// TIA Portal V20 export
FUNCTION_BLOCK "OM_PRM_Access"   // FB82, LAD
{ S7_Optimized_Access := 'TRUE' }
// stored: MemoryReserve 100, SetENOAutomatically false
   VAR_INPUT
      Inputdata_RW_Drv2PLC : "AZ_PrmRW_Drv2PLC";
      ReadParameterID : Word;
      WriteParameterID : Word;
      WriteData : DWord;
      "WR-REQ" : Bool;
   END_VAR
   VAR_OUTPUT
      Outputdata_RW_PLC2Drv : "AZ_PrmRW_PLC2Drv";
      ReadParameterID_R : Word;
      WriteParameterID_R : Word;
      ReadData : DWord;
      "WR-SET-ERR" : Bool;
      "WR-IF-ERR" : Bool;
      "WR-NV-ERR" : Bool;
      "WR-EXE-ERR" : Bool;
      "WR-ERR" : Bool;
      "RD-ERR" : Bool;
      "WR-END" : Bool;
      "SYS-BSY" : Bool;
   END_VAR
BEGIN

REGION Network 1
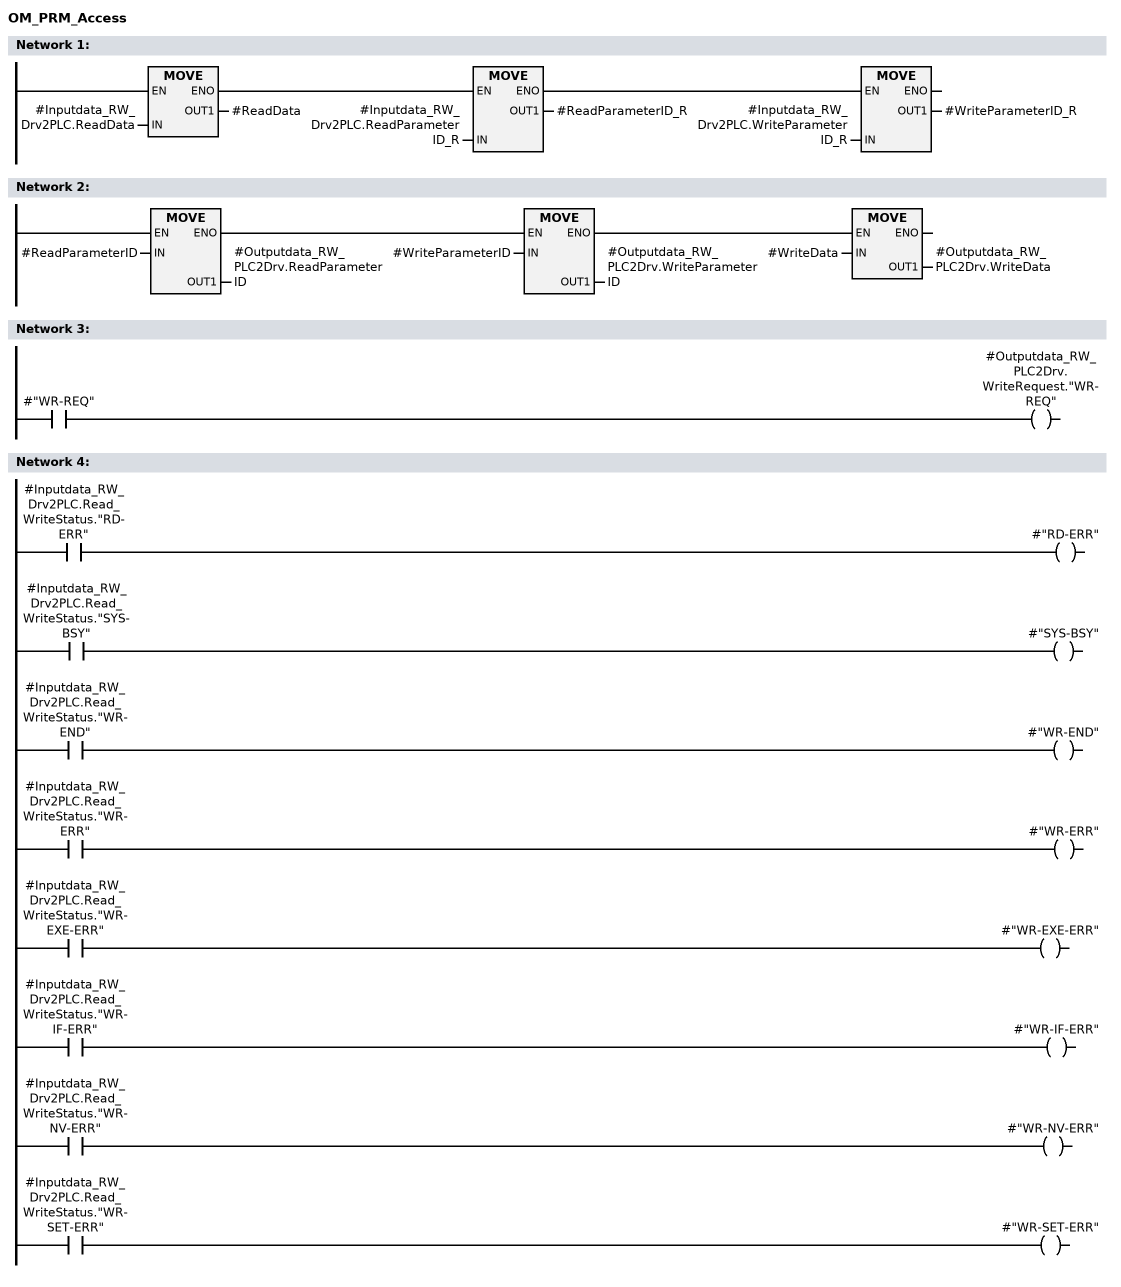
   RUNG wire#powerrail
      Move(in := #Inputdata_RW_Drv2PLC.ReadData, out1 => #ReadData)
      Move(in := #Inputdata_RW_Drv2PLC.ReadParameterID_R, out1 => #ReadParameterID_R)
      Move(in := #Inputdata_RW_Drv2PLC.WriteParameterID_R, out1 => #WriteParameterID_R)
   END_RUNG
   // the same network as SCL:
   #ReadData := #Inputdata_RW_Drv2PLC.ReadData;
   #ReadParameterID_R := #Inputdata_RW_Drv2PLC.ReadParameterID_R;
   #WriteParameterID_R := #Inputdata_RW_Drv2PLC.WriteParameterID_R;
END_REGION

REGION Network 2
   RUNG wire#powerrail
      Move(in := #ReadParameterID, out1 => #Outputdata_RW_PLC2Drv.ReadParameterID)
      Move(in := #WriteParameterID, out1 => #Outputdata_RW_PLC2Drv.WriteParameterID)
      Move(in := #WriteData, out1 => #Outputdata_RW_PLC2Drv.WriteData)
   END_RUNG
   // the same network as SCL:
   #Outputdata_RW_PLC2Drv.ReadParameterID := #ReadParameterID;
   #Outputdata_RW_PLC2Drv.WriteParameterID := #WriteParameterID;
   #Outputdata_RW_PLC2Drv.WriteData := #WriteData;
END_REGION

REGION Network 3
   RUNG wire#powerrail
      Contact( #"WR-REQ" )
      Coil( #Outputdata_RW_PLC2Drv.WriteRequest."WR-REQ" )
   END_RUNG
   // the same network as SCL:
   #Outputdata_RW_PLC2Drv.WriteRequest."WR-REQ" := #"WR-REQ";
END_REGION

REGION Network 4
   RUNG wire#powerrail
      Contact( #Inputdata_RW_Drv2PLC.Read_WriteStatus."RD-ERR" )
      Coil( #"RD-ERR" )
   END_RUNG
   RUNG wire#powerrail
      Contact( #Inputdata_RW_Drv2PLC.Read_WriteStatus."SYS-BSY" )
      Coil( #"SYS-BSY" )
   END_RUNG
   RUNG wire#powerrail
      Contact( #Inputdata_RW_Drv2PLC.Read_WriteStatus."WR-END" )
      Coil( #"WR-END" )
   END_RUNG
   RUNG wire#powerrail
      Contact( #Inputdata_RW_Drv2PLC.Read_WriteStatus."WR-ERR" )
      Coil( #"WR-ERR" )
   END_RUNG
   RUNG wire#powerrail
      Contact( #Inputdata_RW_Drv2PLC.Read_WriteStatus."WR-EXE-ERR" )
      Coil( #"WR-EXE-ERR" )
   END_RUNG
   RUNG wire#powerrail
      Contact( #Inputdata_RW_Drv2PLC.Read_WriteStatus."WR-IF-ERR" )
      Coil( #"WR-IF-ERR" )
   END_RUNG
   RUNG wire#powerrail
      Contact( #Inputdata_RW_Drv2PLC.Read_WriteStatus."WR-NV-ERR" )
      Coil( #"WR-NV-ERR" )
   END_RUNG
   RUNG wire#powerrail
      Contact( #Inputdata_RW_Drv2PLC.Read_WriteStatus."WR-SET-ERR" )
      Coil( #"WR-SET-ERR" )
   END_RUNG
   // the same network as SCL:
   #"RD-ERR" := #Inputdata_RW_Drv2PLC.Read_WriteStatus."RD-ERR";
   #"SYS-BSY" := #Inputdata_RW_Drv2PLC.Read_WriteStatus."SYS-BSY";
   #"WR-END" := #Inputdata_RW_Drv2PLC.Read_WriteStatus."WR-END";
   #"WR-ERR" := #Inputdata_RW_Drv2PLC.Read_WriteStatus."WR-ERR";
   #"WR-EXE-ERR" := #Inputdata_RW_Drv2PLC.Read_WriteStatus."WR-EXE-ERR";
   #"WR-IF-ERR" := #Inputdata_RW_Drv2PLC.Read_WriteStatus."WR-IF-ERR";
   #"WR-NV-ERR" := #Inputdata_RW_Drv2PLC.Read_WriteStatus."WR-NV-ERR";
   #"WR-SET-ERR" := #Inputdata_RW_Drv2PLC.Read_WriteStatus."WR-SET-ERR";
END_REGION
END_FUNCTION_BLOCK
